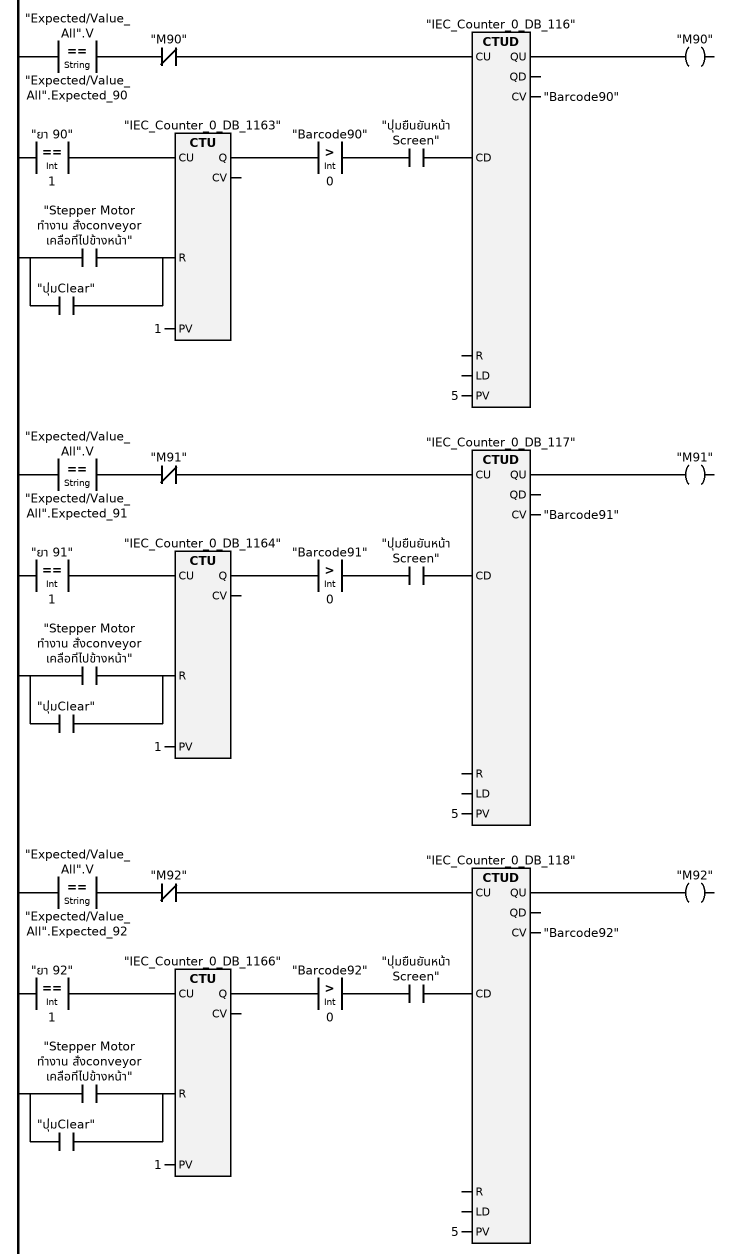
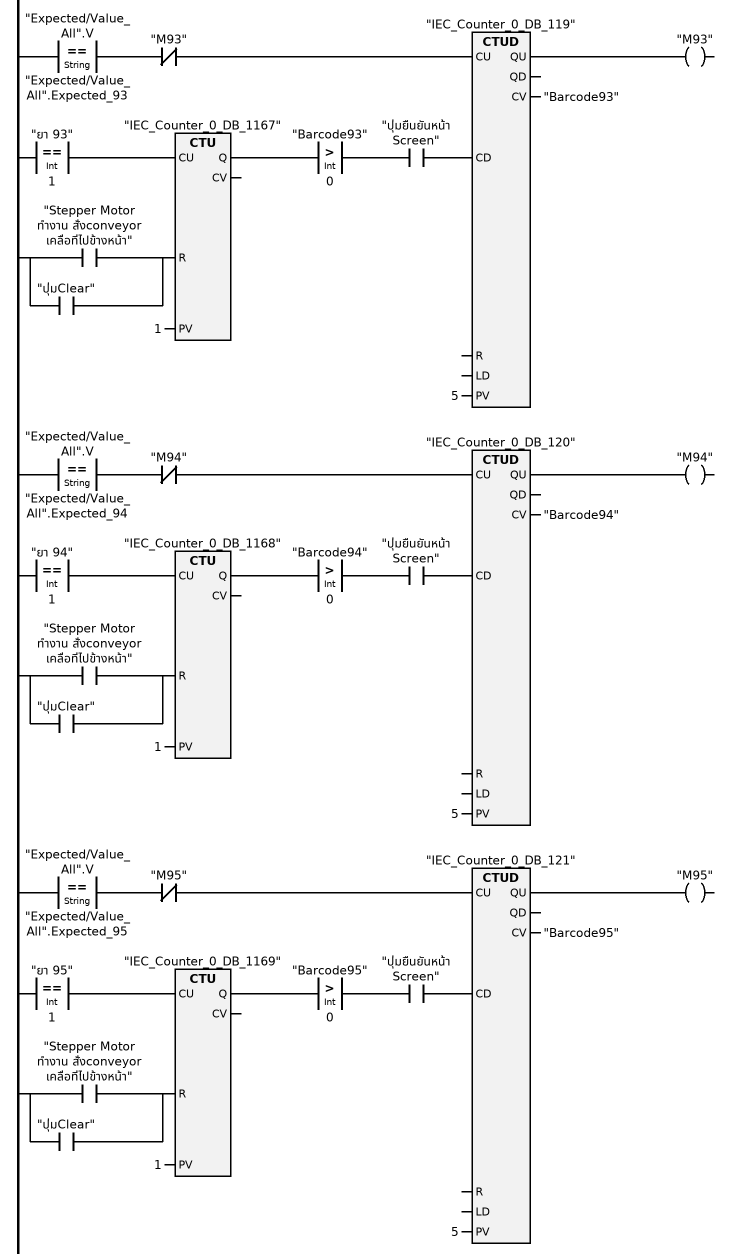
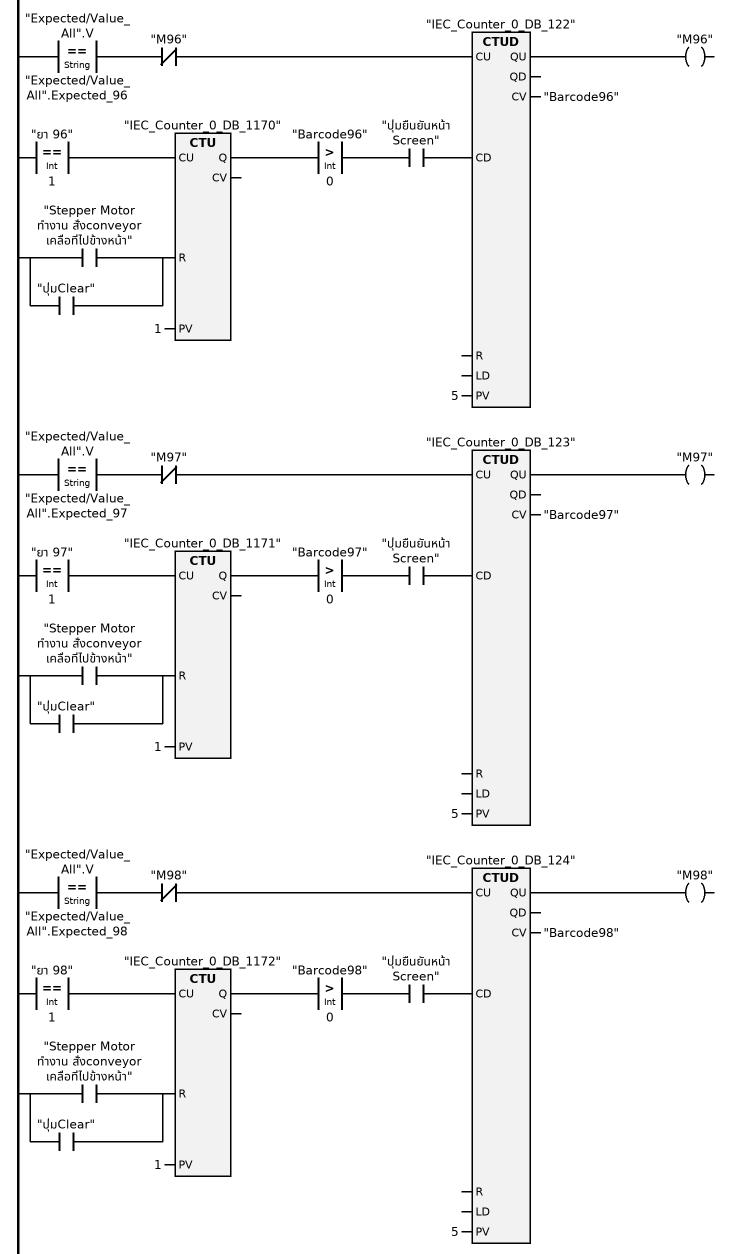
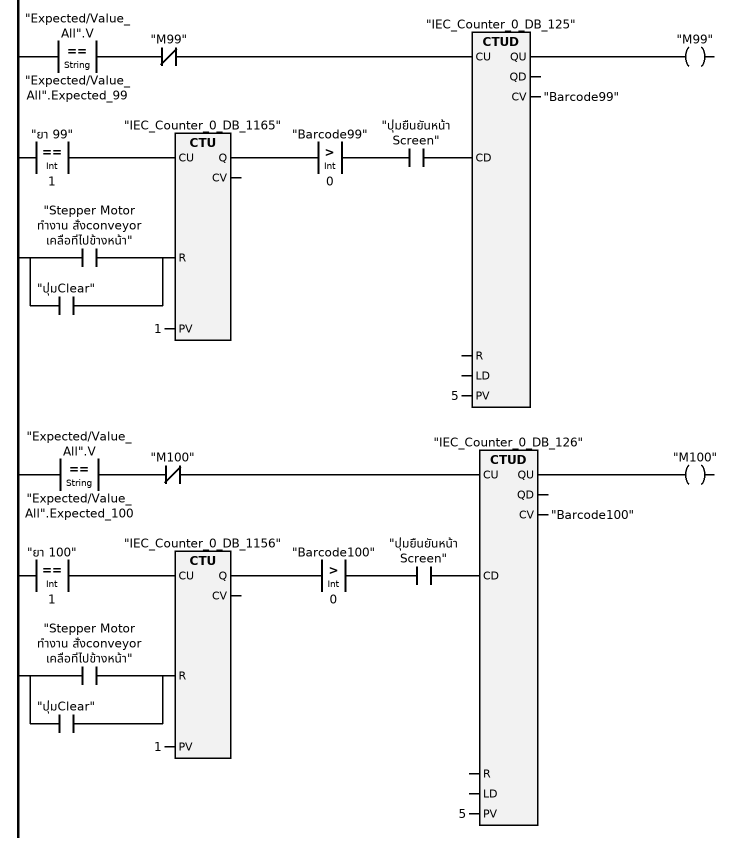
   "IEC_Counter_0_DB_1153".CTU(CU := "ยา 81" = 1,
                           R := "Stepper Motor ทำงาน สั่งconveyor เคลื่อที่ไปข้างหน้า" OR "ปุ่มClear",
                           PV := 1);
   "IEC_Counter_0_DB_107".CTUD(CU := ("Expected/Value_All".V = "Expected/Value_All".Expected_81) AND NOT "M81",
                           CD := "IEC_Counter_0_DB_1153".Q AND ("Barcode81" > 0) AND "ปุ่มยืนยันหน้า Screen",
                           PV := 5,
                           CV => "Barcode81");
   "M81" := "IEC_Counter_0_DB_107".QU;
   "IEC_Counter_0_DB_1154".CTU(CU := "ยา 82" = 1,
                           R := "Stepper Motor ทำงาน สั่งconveyor เคลื่อที่ไปข้างหน้า" OR "ปุ่มClear",
                           PV := 1);
   "IEC_Counter_0_DB_108".CTUD(CU := ("Expected/Value_All".V = "Expected/Value_All".Expected_82) AND NOT "M82",
                           CD := "IEC_Counter_0_DB_1154".Q AND ("Barcode82" > 0) AND "ปุ่มยืนยันหน้า Screen",
                           PV := 5,
                           CV => "Barcode82");
   "M82" := "IEC_Counter_0_DB_108".QU;
   "IEC_Counter_0_DB_1155".CTU(CU := "ยา 83" = 1,
                           R := "Stepper Motor ทำงาน สั่งconveyor เคลื่อที่ไปข้างหน้า" OR "ปุ่มClear",
                           PV := 1);
   "IEC_Counter_0_DB_109".CTUD(CU := ("Expected/Value_All".V = "Expected/Value_All".Expected_83) AND NOT "M83",
                           CD := "IEC_Counter_0_DB_1155".Q AND ("Barcode83" > 0) AND "ปุ่มยืนยันหน้า Screen",
                           PV := 5,
                           CV => "Barcode83");
   "M83" := "IEC_Counter_0_DB_109".QU;
   "IEC_Counter_0_DB_1157".CTU(CU := "ยา 84" = 1,
                           R := "Stepper Motor ทำงาน สั่งconveyor เคลื่อที่ไปข้างหน้า" OR "ปุ่มClear",
                           PV := 1);
   "IEC_Counter_0_DB_110".CTUD(CU := ("Expected/Value_All".V = "Expected/Value_All".Expected_84) AND NOT "M84",
                           CD := "IEC_Counter_0_DB_1157".Q AND ("Barcode84" > 0) AND "ปุ่มยืนยันหน้า Screen",
                           PV := 5,
                           CV => "Barcode84");
   "M84" := "IEC_Counter_0_DB_110".QU;
   "IEC_Counter_0_DB_1158".CTU(CU := "ยา 85" = 1,
                           R := "Stepper Motor ทำงาน สั่งconveyor เคลื่อที่ไปข้างหน้า" OR "ปุ่มClear",
                           PV := 1);
   "IEC_Counter_0_DB_111".CTUD(CU := ("Expected/Value_All".V = "Expected/Value_All".Expected_85) AND NOT "M85",
                           CD := "IEC_Counter_0_DB_1158".Q AND ("Barcode85" > 0) AND "ปุ่มยืนยันหน้า Screen",
                           PV := 5,
                           CV => "Barcode85");
   "M85" := "IEC_Counter_0_DB_111".QU;
   "IEC_Counter_0_DB_1159".CTU(CU := "ยา 86" = 1,
                           R := "Stepper Motor ทำงาน สั่งconveyor เคลื่อที่ไปข้างหน้า" OR "ปุ่มClear",
                           PV := 1);
   "IEC_Counter_0_DB_112".CTUD(CU := ("Expected/Value_All".V = "Expected/Value_All".Expected_86) AND NOT "M86",
                           CD := "IEC_Counter_0_DB_1159".Q AND ("Barcode86" > 0) AND "ปุ่มยืนยันหน้า Screen",
                           PV := 5,
                           CV => "Barcode86");
   "M86" := "IEC_Counter_0_DB_112".QU;
   "IEC_Counter_0_DB_1160".CTU(CU := "ยา 87" = 1,
                           R := "Stepper Motor ทำงาน สั่งconveyor เคลื่อที่ไปข้างหน้า" OR "ปุ่มClear",
                           PV := 1);
   "IEC_Counter_0_DB_113".CTUD(CU := ("Expected/Value_All".V = "Expected/Value_All".Expected_87) AND NOT "M87",
                           CD := "IEC_Counter_0_DB_1160".Q AND ("Barcode87" > 0) AND "ปุ่มยืนยันหน้า Screen",
                           PV := 5,
                           CV => "Barcode87");
   "M87" := "IEC_Counter_0_DB_113".QU;
   "IEC_Counter_0_DB_1161".CTU(CU := "ยา 88" = 1,
                           R := "Stepper Motor ทำงาน สั่งconveyor เคลื่อที่ไปข้างหน้า" OR "ปุ่มClear",
                           PV := 1);
   "IEC_Counter_0_DB_114".CTUD(CU := ("Expected/Value_All".V = "Expected/Value_All".Expected_88) AND NOT "M88",
                           CD := "IEC_Counter_0_DB_1161".Q AND ("Barcode88" > 0) AND "ปุ่มยืนยันหน้า Screen",
                           PV := 5,
                           CV => "Barcode88");
   "M88" := "IEC_Counter_0_DB_114".QU;
   "IEC_Counter_0_DB_1162".CTU(CU := "ยา 89" = 1,
                           R := "Stepper Motor ทำงาน สั่งconveyor เคลื่อที่ไปข้างหน้า" OR "ปุ่มClear",
                           PV := 1);
   "IEC_Counter_0_DB_115".CTUD(CU := ("Expected/Value_All".V = "Expected/Value_All".Expected_89) AND NOT "M89",
                           CD := "IEC_Counter_0_DB_1162".Q AND ("Barcode89" > 0) AND "ปุ่มยืนยันหน้า Screen",
                           PV := 5,
                           CV => "Barcode89");
   "M89" := "IEC_Counter_0_DB_115".QU;
   "IEC_Counter_0_DB_1163".CTU(CU := "ยา 90" = 1,
                           R := "Stepper Motor ทำงาน สั่งconveyor เคลื่อที่ไปข้างหน้า" OR "ปุ่มClear",
                           PV := 1);
   "IEC_Counter_0_DB_116".CTUD(CU := ("Expected/Value_All".V = "Expected/Value_All".Expected_90) AND NOT "M90",
                           CD := "IEC_Counter_0_DB_1163".Q AND ("Barcode90" > 0) AND "ปุ่มยืนยันหน้า Screen",
                           PV := 5,
                           CV => "Barcode90");
   "M90" := "IEC_Counter_0_DB_116".QU;
   "IEC_Counter_0_DB_1164".CTU(CU := "ยา 91" = 1,
                           R := "Stepper Motor ทำงาน สั่งconveyor เคลื่อที่ไปข้างหน้า" OR "ปุ่มClear",
                           PV := 1);
   "IEC_Counter_0_DB_117".CTUD(CU := ("Expected/Value_All".V = "Expected/Value_All".Expected_91) AND NOT "M91",
                           CD := "IEC_Counter_0_DB_1164".Q AND ("Barcode91" > 0) AND "ปุ่มยืนยันหน้า Screen",
                           PV := 5,
                           CV => "Barcode91");
   "M91" := "IEC_Counter_0_DB_117".QU;
   "IEC_Counter_0_DB_1166".CTU(CU := "ยา 92" = 1,
                           R := "Stepper Motor ทำงาน สั่งconveyor เคลื่อที่ไปข้างหน้า" OR "ปุ่มClear",
                           PV := 1);
   "IEC_Counter_0_DB_118".CTUD(CU := ("Expected/Value_All".V = "Expected/Value_All".Expected_92) AND NOT "M92",
                           CD := "IEC_Counter_0_DB_1166".Q AND ("Barcode92" > 0) AND "ปุ่มยืนยันหน้า Screen",
                           PV := 5,
                           CV => "Barcode92");
   "M92" := "IEC_Counter_0_DB_118".QU;
   "IEC_Counter_0_DB_1167".CTU(CU := "ยา 93" = 1,
                           R := "Stepper Motor ทำงาน สั่งconveyor เคลื่อที่ไปข้างหน้า" OR "ปุ่มClear",
                           PV := 1);
   "IEC_Counter_0_DB_119".CTUD(CU := ("Expected/Value_All".V = "Expected/Value_All".Expected_93) AND NOT "M93",
                           CD := "IEC_Counter_0_DB_1167".Q AND ("Barcode93" > 0) AND "ปุ่มยืนยันหน้า Screen",
                           PV := 5,
                           CV => "Barcode93");
   "M93" := "IEC_Counter_0_DB_119".QU;
   "IEC_Counter_0_DB_1168".CTU(CU := "ยา 94" = 1,
                           R := "Stepper Motor ทำงาน สั่งconveyor เคลื่อที่ไปข้างหน้า" OR "ปุ่มClear",
                           PV := 1);
   "IEC_Counter_0_DB_120".CTUD(CU := ("Expected/Value_All".V = "Expected/Value_All".Expected_94) AND NOT "M94",
                           CD := "IEC_Counter_0_DB_1168".Q AND ("Barcode94" > 0) AND "ปุ่มยืนยันหน้า Screen",
                           PV := 5,
                           CV => "Barcode94");
   "M94" := "IEC_Counter_0_DB_120".QU;
   "IEC_Counter_0_DB_1169".CTU(CU := "ยา 95" = 1,
                           R := "Stepper Motor ทำงาน สั่งconveyor เคลื่อที่ไปข้างหน้า" OR "ปุ่มClear",
                           PV := 1);
   "IEC_Counter_0_DB_121".CTUD(CU := ("Expected/Value_All".V = "Expected/Value_All".Expected_95) AND NOT "M95",
                           CD := "IEC_Counter_0_DB_1169".Q AND ("Barcode95" > 0) AND "ปุ่มยืนยันหน้า Screen",
                           PV := 5,
                           CV => "Barcode95");
   "M95" := "IEC_Counter_0_DB_121".QU;
   "IEC_Counter_0_DB_1170".CTU(CU := "ยา 96" = 1,
                           R := "Stepper Motor ทำงาน สั่งconveyor เคลื่อที่ไปข้างหน้า" OR "ปุ่มClear",
                           PV := 1);
   "IEC_Counter_0_DB_122".CTUD(CU := ("Expected/Value_All".V = "Expected/Value_All".Expected_96) AND NOT "M96",
                           CD := "IEC_Counter_0_DB_1170".Q AND ("Barcode96" > 0) AND "ปุ่มยืนยันหน้า Screen",
                           PV := 5,
                           CV => "Barcode96");
   "M96" := "IEC_Counter_0_DB_122".QU;
   "IEC_Counter_0_DB_1171".CTU(CU := "ยา 97" = 1,
                           R := "Stepper Motor ทำงาน สั่งconveyor เคลื่อที่ไปข้างหน้า" OR "ปุ่มClear",
                           PV := 1);
   "IEC_Counter_0_DB_123".CTUD(CU := ("Expected/Value_All".V = "Expected/Value_All".Expected_97) AND NOT "M97",
                           CD := "IEC_Counter_0_DB_1171".Q AND ("Barcode97" > 0) AND "ปุ่มยืนยันหน้า Screen",
                           PV := 5,
                           CV => "Barcode97");
   "M97" := "IEC_Counter_0_DB_123".QU;
   "IEC_Counter_0_DB_1172".CTU(CU := "ยา 98" = 1,
                           R := "Stepper Motor ทำงาน สั่งconveyor เคลื่อที่ไปข้างหน้า" OR "ปุ่มClear",
                           PV := 1);
   "IEC_Counter_0_DB_124".CTUD(CU := ("Expected/Value_All".V = "Expected/Value_All".Expected_98) AND NOT "M98",
                           CD := "IEC_Counter_0_DB_1172".Q AND ("Barcode98" > 0) AND "ปุ่มยืนยันหน้า Screen",
                           PV := 5,
                           CV => "Barcode98");
   "M98" := "IEC_Counter_0_DB_124".QU;
   "IEC_Counter_0_DB_1165".CTU(CU := "ยา 99" = 1,
                           R := "Stepper Motor ทำงาน สั่งconveyor เคลื่อที่ไปข้างหน้า" OR "ปุ่มClear",
                           PV := 1);
   "IEC_Counter_0_DB_125".CTUD(CU := ("Expected/Value_All".V = "Expected/Value_All".Expected_99) AND NOT "M99",
                           CD := "IEC_Counter_0_DB_1165".Q AND ("Barcode99" > 0) AND "ปุ่มยืนยันหน้า Screen",
                           PV := 5,
                           CV => "Barcode99");
   "M99" := "IEC_Counter_0_DB_125".QU;
   "IEC_Counter_0_DB_1156".CTU(CU := "ยา 100" = 1,
                           R := "Stepper Motor ทำงาน สั่งconveyor เคลื่อที่ไปข้างหน้า" OR "ปุ่มClear",
                           PV := 1);
   "IEC_Counter_0_DB_126".CTUD(CU := ("Expected/Value_All".V = "Expected/Value_All".Expected_100) AND NOT "M100",
                           CD := "IEC_Counter_0_DB_1156".Q AND ("Barcode100" > 0) AND "ปุ่มยืนยันหน้า Screen",
                           PV := 5,
                           CV => "Barcode100");
   "M100" := "IEC_Counter_0_DB_126".QU;
END_REGION

REGION Network 6
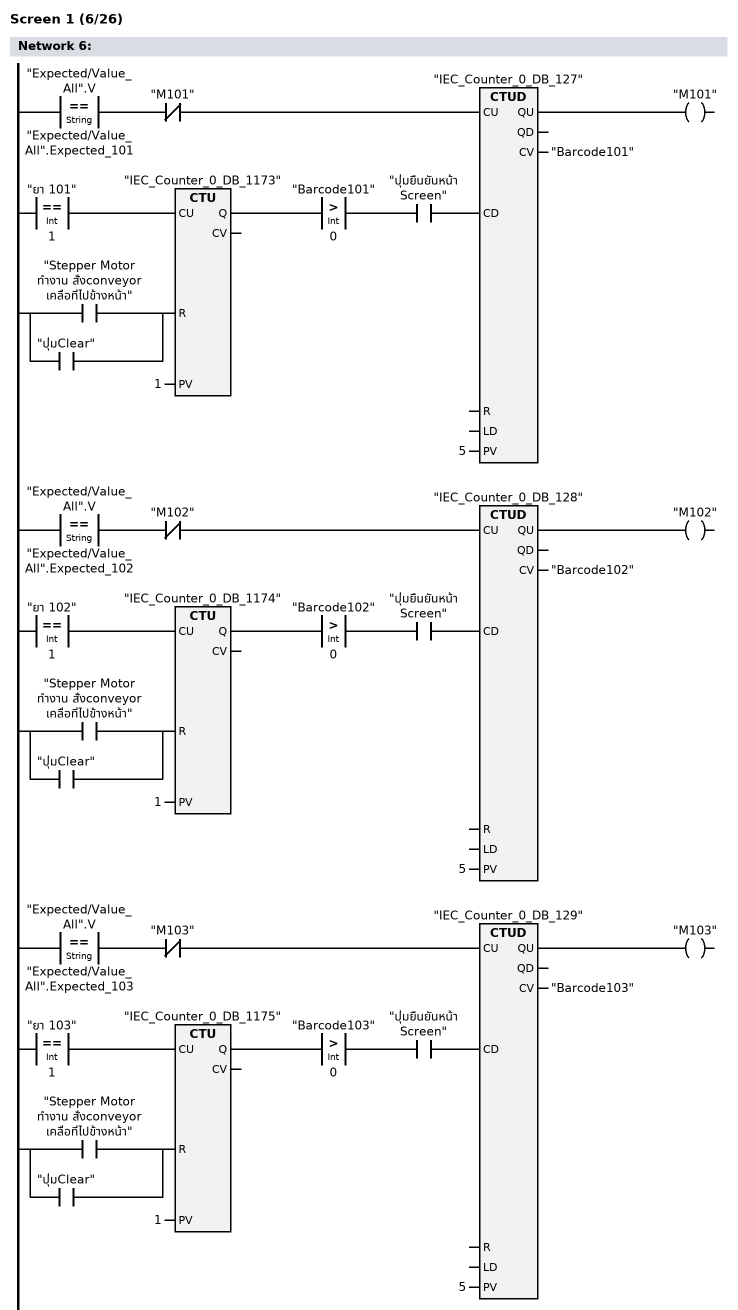
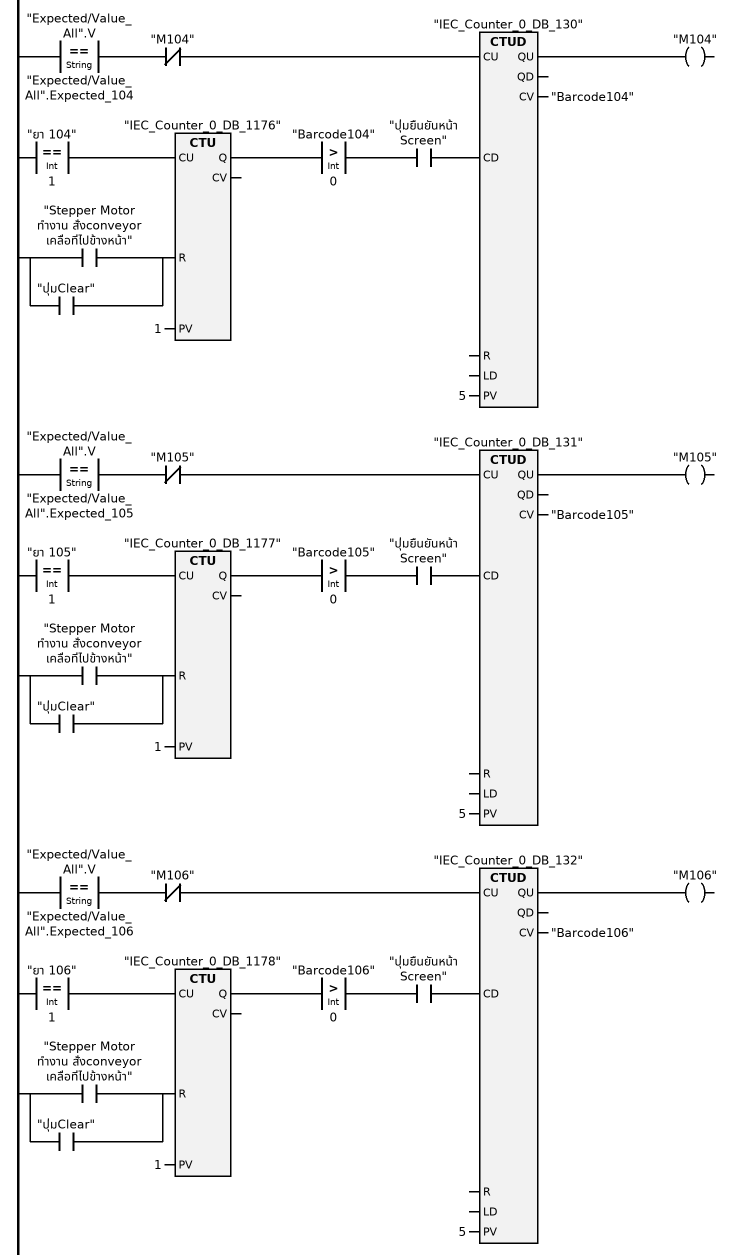
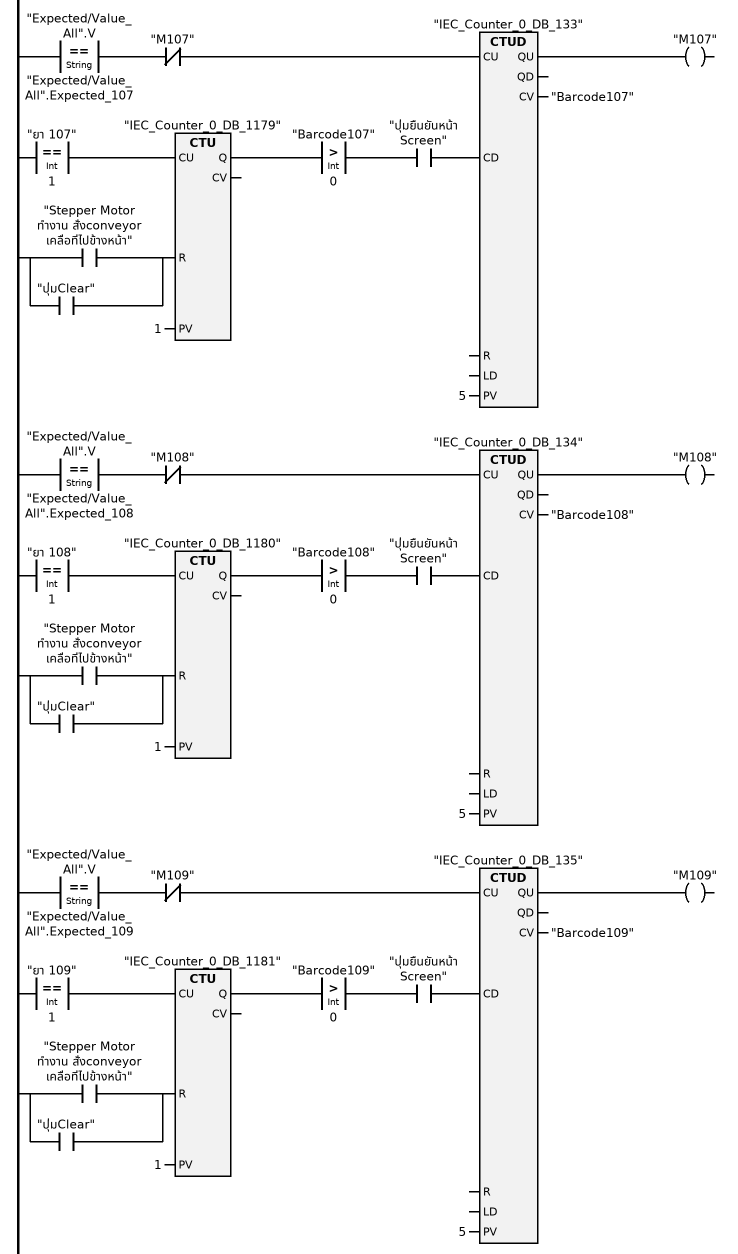
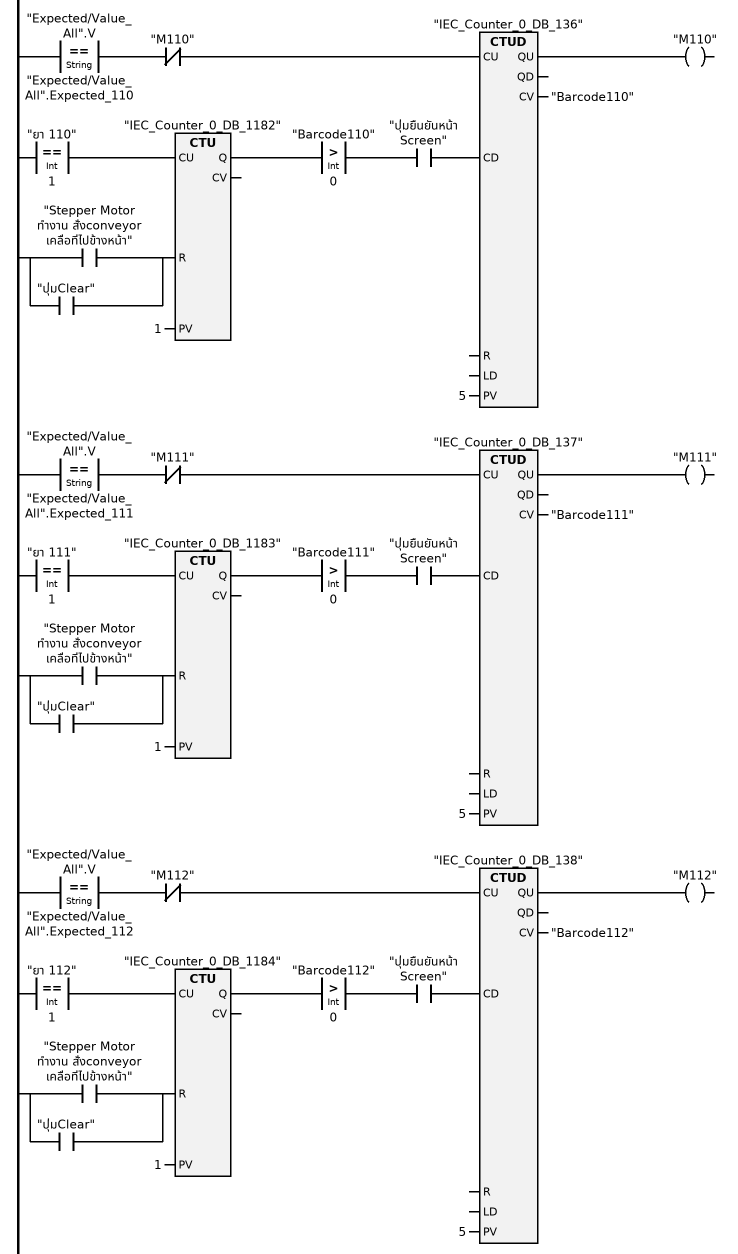
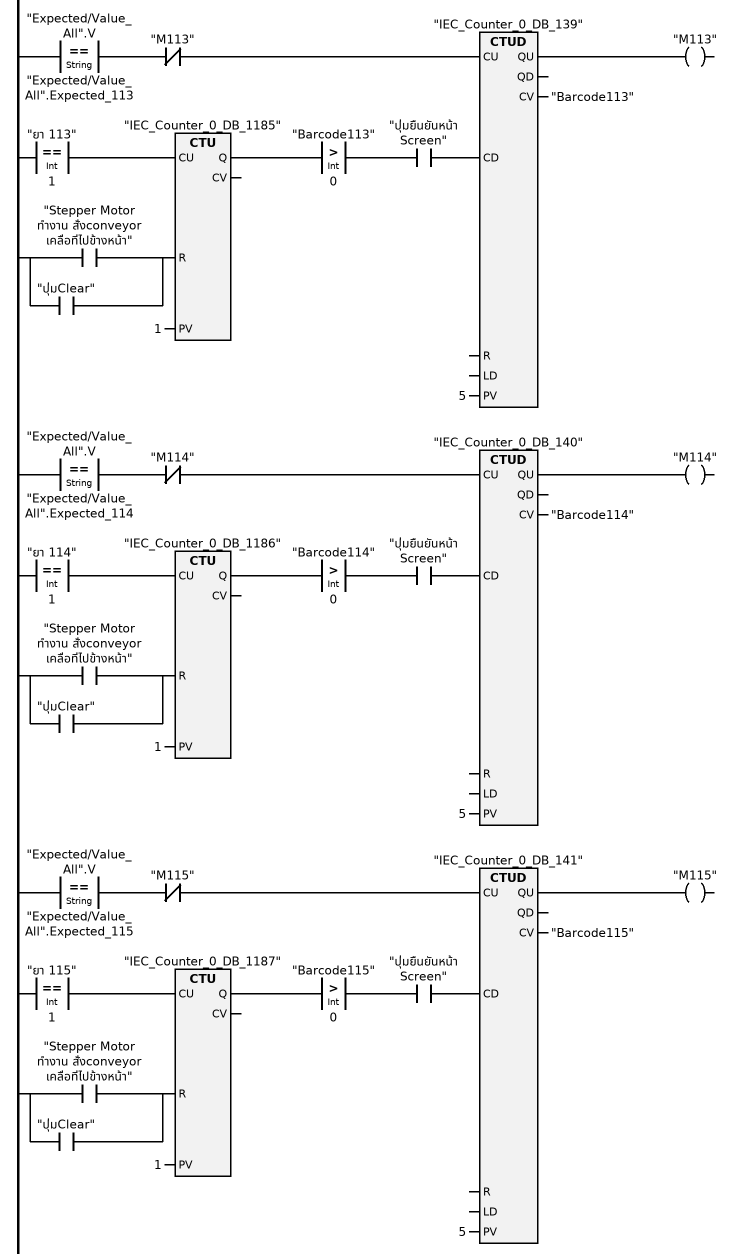
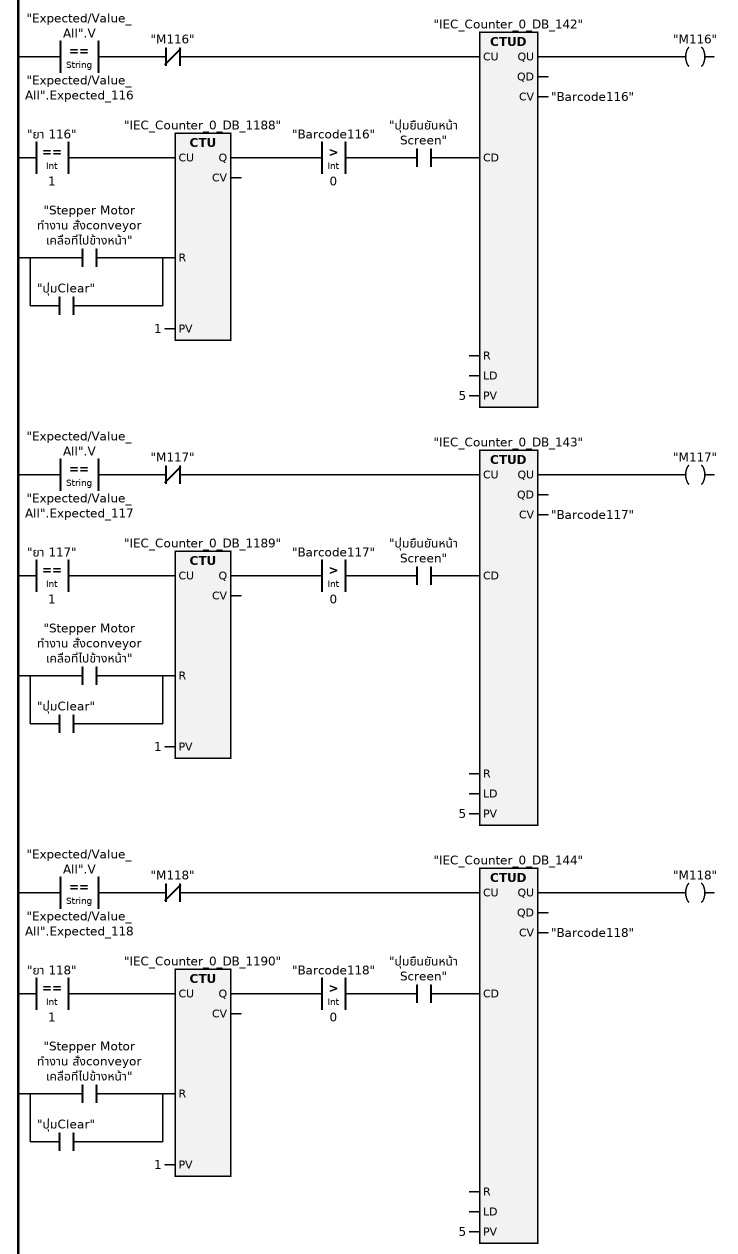
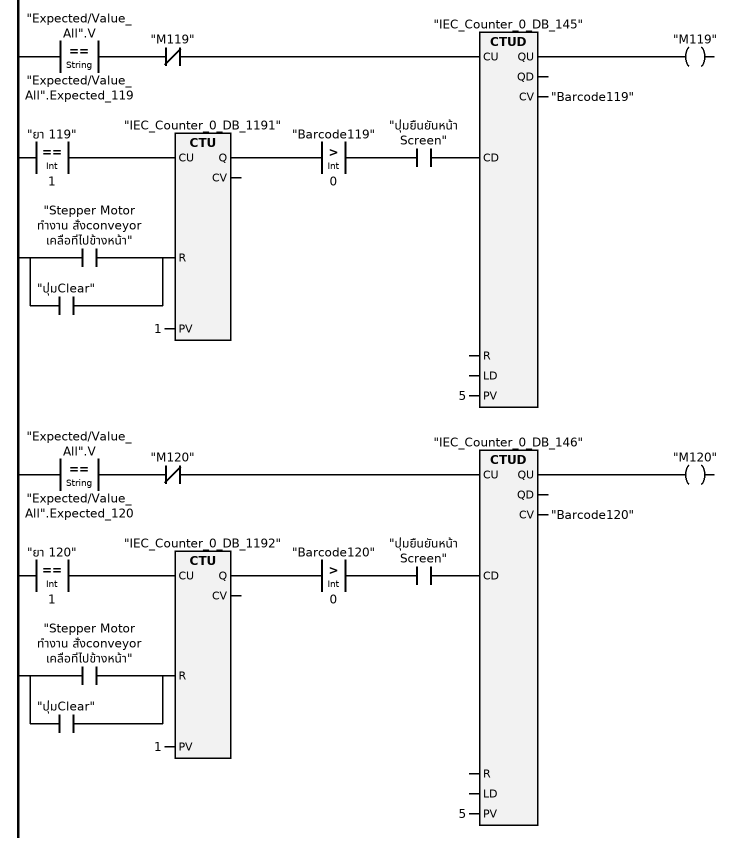
   "IEC_Counter_0_DB_1173".CTU(CU := "ยา 101" = 1,
                           R := "Stepper Motor ทำงาน สั่งconveyor เคลื่อที่ไปข้างหน้า" OR "ปุ่มClear",
                           PV := 1);
   "IEC_Counter_0_DB_127".CTUD(CU := ("Expected/Value_All".V = "Expected/Value_All".Expected_101) AND NOT "M101",
                           CD := "IEC_Counter_0_DB_1173".Q AND ("Barcode101" > 0) AND "ปุ่มยืนยันหน้า Screen",
                           PV := 5,
                           CV => "Barcode101");
   "M101" := "IEC_Counter_0_DB_127".QU;
   "IEC_Counter_0_DB_1174".CTU(CU := "ยา 102" = 1,
                           R := "Stepper Motor ทำงาน สั่งconveyor เคลื่อที่ไปข้างหน้า" OR "ปุ่มClear",
                           PV := 1);
   "IEC_Counter_0_DB_128".CTUD(CU := ("Expected/Value_All".V = "Expected/Value_All".Expected_102) AND NOT "M102",
                           CD := "IEC_Counter_0_DB_1174".Q AND ("Barcode102" > 0) AND "ปุ่มยืนยันหน้า Screen",
                           PV := 5,
                           CV => "Barcode102");
   "M102" := "IEC_Counter_0_DB_128".QU;
   "IEC_Counter_0_DB_1175".CTU(CU := "ยา 103" = 1,
                           R := "Stepper Motor ทำงาน สั่งconveyor เคลื่อที่ไปข้างหน้า" OR "ปุ่มClear",
                           PV := 1);
   "IEC_Counter_0_DB_129".CTUD(CU := ("Expected/Value_All".V = "Expected/Value_All".Expected_103) AND NOT "M103",
                           CD := "IEC_Counter_0_DB_1175".Q AND ("Barcode103" > 0) AND "ปุ่มยืนยันหน้า Screen",
                           PV := 5,
                           CV => "Barcode103");
   "M103" := "IEC_Counter_0_DB_129".QU;
   "IEC_Counter_0_DB_1176".CTU(CU := "ยา 104" = 1,
                           R := "Stepper Motor ทำงาน สั่งconveyor เคลื่อที่ไปข้างหน้า" OR "ปุ่มClear",
                           PV := 1);
   "IEC_Counter_0_DB_130".CTUD(CU := ("Expected/Value_All".V = "Expected/Value_All".Expected_104) AND NOT "M104",
                           CD := "IEC_Counter_0_DB_1176".Q AND ("Barcode104" > 0) AND "ปุ่มยืนยันหน้า Screen",
                           PV := 5,
                           CV => "Barcode104");
   "M104" := "IEC_Counter_0_DB_130".QU;
   "IEC_Counter_0_DB_1177".CTU(CU := "ยา 105" = 1,
                           R := "Stepper Motor ทำงาน สั่งconveyor เคลื่อที่ไปข้างหน้า" OR "ปุ่มClear",
                           PV := 1);
   "IEC_Counter_0_DB_131".CTUD(CU := ("Expected/Value_All".V = "Expected/Value_All".Expected_105) AND NOT "M105",
                           CD := "IEC_Counter_0_DB_1177".Q AND ("Barcode105" > 0) AND "ปุ่มยืนยันหน้า Screen",
                           PV := 5,
                           CV => "Barcode105");
   "M105" := "IEC_Counter_0_DB_131".QU;
   "IEC_Counter_0_DB_1178".CTU(CU := "ยา 106" = 1,
                           R := "Stepper Motor ทำงาน สั่งconveyor เคลื่อที่ไปข้างหน้า" OR "ปุ่มClear",
                           PV := 1);
   "IEC_Counter_0_DB_132".CTUD(CU := ("Expected/Value_All".V = "Expected/Value_All".Expected_106) AND NOT "M106",
                           CD := "IEC_Counter_0_DB_1178".Q AND ("Barcode106" > 0) AND "ปุ่มยืนยันหน้า Screen",
                           PV := 5,
                           CV => "Barcode106");
   "M106" := "IEC_Counter_0_DB_132".QU;
   "IEC_Counter_0_DB_1179".CTU(CU := "ยา 107" = 1,
                           R := "Stepper Motor ทำงาน สั่งconveyor เคลื่อที่ไปข้างหน้า" OR "ปุ่มClear",
                           PV := 1);
   "IEC_Counter_0_DB_133".CTUD(CU := ("Expected/Value_All".V = "Expected/Value_All".Expected_107) AND NOT "M107",
                           CD := "IEC_Counter_0_DB_1179".Q AND ("Barcode107" > 0) AND "ปุ่มยืนยันหน้า Screen",
                           PV := 5,
                           CV => "Barcode107");
   "M107" := "IEC_Counter_0_DB_133".QU;
   "IEC_Counter_0_DB_1180".CTU(CU := "ยา 108" = 1,
                           R := "Stepper Motor ทำงาน สั่งconveyor เคลื่อที่ไปข้างหน้า" OR "ปุ่มClear",
                           PV := 1);
   "IEC_Counter_0_DB_134".CTUD(CU := ("Expected/Value_All".V = "Expected/Value_All".Expected_108) AND NOT "M108",
                           CD := "IEC_Counter_0_DB_1180".Q AND ("Barcode108" > 0) AND "ปุ่มยืนยันหน้า Screen",
                           PV := 5,
                           CV => "Barcode108");
   "M108" := "IEC_Counter_0_DB_134".QU;
   "IEC_Counter_0_DB_1181".CTU(CU := "ยา 109" = 1,
                           R := "Stepper Motor ทำงาน สั่งconveyor เคลื่อที่ไปข้างหน้า" OR "ปุ่มClear",
                           PV := 1);
   "IEC_Counter_0_DB_135".CTUD(CU := ("Expected/Value_All".V = "Expected/Value_All".Expected_109) AND NOT "M109",
                           CD := "IEC_Counter_0_DB_1181".Q AND ("Barcode109" > 0) AND "ปุ่มยืนยันหน้า Screen",
                           PV := 5,
                           CV => "Barcode109");
   "M109" := "IEC_Counter_0_DB_135".QU;
   "IEC_Counter_0_DB_1182".CTU(CU := "ยา 110" = 1,
                           R := "Stepper Motor ทำงาน สั่งconveyor เคลื่อที่ไปข้างหน้า" OR "ปุ่มClear",
                           PV := 1);
   "IEC_Counter_0_DB_136".CTUD(CU := ("Expected/Value_All".V = "Expected/Value_All".Expected_110) AND NOT "M110",
                           CD := "IEC_Counter_0_DB_1182".Q AND ("Barcode110" > 0) AND "ปุ่มยืนยันหน้า Screen",
                           PV := 5,
                           CV => "Barcode110");
   "M110" := "IEC_Counter_0_DB_136".QU;
   "IEC_Counter_0_DB_1183".CTU(CU := "ยา 111" = 1,
                           R := "Stepper Motor ทำงาน สั่งconveyor เคลื่อที่ไปข้างหน้า" OR "ปุ่มClear",
                           PV := 1);
   "IEC_Counter_0_DB_137".CTUD(CU := ("Expected/Value_All".V = "Expected/Value_All".Expected_111) AND NOT "M111",
                           CD := "IEC_Counter_0_DB_1183".Q AND ("Barcode111" > 0) AND "ปุ่มยืนยันหน้า Screen",
                           PV := 5,
                           CV => "Barcode111");
   "M111" := "IEC_Counter_0_DB_137".QU;
   "IEC_Counter_0_DB_1184".CTU(CU := "ยา 112" = 1,
                           R := "Stepper Motor ทำงาน สั่งconveyor เคลื่อที่ไปข้างหน้า" OR "ปุ่มClear",
                           PV := 1);
   "IEC_Counter_0_DB_138".CTUD(CU := ("Expected/Value_All".V = "Expected/Value_All".Expected_112) AND NOT "M112",
                           CD := "IEC_Counter_0_DB_1184".Q AND ("Barcode112" > 0) AND "ปุ่มยืนยันหน้า Screen",
                           PV := 5,
                           CV => "Barcode112");
   "M112" := "IEC_Counter_0_DB_138".QU;
   "IEC_Counter_0_DB_1185".CTU(CU := "ยา 113" = 1,
                           R := "Stepper Motor ทำงาน สั่งconveyor เคลื่อที่ไปข้างหน้า" OR "ปุ่มClear",
                           PV := 1);
   "IEC_Counter_0_DB_139".CTUD(CU := ("Expected/Value_All".V = "Expected/Value_All".Expected_113) AND NOT "M113",
                           CD := "IEC_Counter_0_DB_1185".Q AND ("Barcode113" > 0) AND "ปุ่มยืนยันหน้า Screen",
                           PV := 5,
                           CV => "Barcode113");
   "M113" := "IEC_Counter_0_DB_139".QU;
   "IEC_Counter_0_DB_1186".CTU(CU := "ยา 114" = 1,
                           R := "Stepper Motor ทำงาน สั่งconveyor เคลื่อที่ไปข้างหน้า" OR "ปุ่มClear",
                           PV := 1);
   "IEC_Counter_0_DB_140".CTUD(CU := ("Expected/Value_All".V = "Expected/Value_All".Expected_114) AND NOT "M114",
                           CD := "IEC_Counter_0_DB_1186".Q AND ("Barcode114" > 0) AND "ปุ่มยืนยันหน้า Screen",
                           PV := 5,
                           CV => "Barcode114");
   "M114" := "IEC_Counter_0_DB_140".QU;
   "IEC_Counter_0_DB_1187".CTU(CU := "ยา 115" = 1,
                           R := "Stepper Motor ทำงาน สั่งconveyor เคลื่อที่ไปข้างหน้า" OR "ปุ่มClear",
                           PV := 1);
   "IEC_Counter_0_DB_141".CTUD(CU := ("Expected/Value_All".V = "Expected/Value_All".Expected_115) AND NOT "M115",
                           CD := "IEC_Counter_0_DB_1187".Q AND ("Barcode115" > 0) AND "ปุ่มยืนยันหน้า Screen",
                           PV := 5,
                           CV => "Barcode115");
   "M115" := "IEC_Counter_0_DB_141".QU;
   "IEC_Counter_0_DB_1188".CTU(CU := "ยา 116" = 1,
                           R := "Stepper Motor ทำงาน สั่งconveyor เคลื่อที่ไปข้างหน้า" OR "ปุ่มClear",
                           PV := 1);
   "IEC_Counter_0_DB_142".CTUD(CU := ("Expected/Value_All".V = "Expected/Value_All".Expected_116) AND NOT "M116",
                           CD := "IEC_Counter_0_DB_1188".Q AND ("Barcode116" > 0) AND "ปุ่มยืนยันหน้า Screen",
                           PV := 5,
                           CV => "Barcode116");
   "M116" := "IEC_Counter_0_DB_142".QU;
   "IEC_Counter_0_DB_1189".CTU(CU := "ยา 117" = 1,
                           R := "Stepper Motor ทำงาน สั่งconveyor เคลื่อที่ไปข้างหน้า" OR "ปุ่มClear",
                           PV := 1);
   "IEC_Counter_0_DB_143".CTUD(CU := ("Expected/Value_All".V = "Expected/Value_All".Expected_117) AND NOT "M117",
                           CD := "IEC_Counter_0_DB_1189".Q AND ("Barcode117" > 0) AND "ปุ่มยืนยันหน้า Screen",
                           PV := 5,
                           CV => "Barcode117");
   "M117" := "IEC_Counter_0_DB_143".QU;
   "IEC_Counter_0_DB_1190".CTU(CU := "ยา 118" = 1,
                           R := "Stepper Motor ทำงาน สั่งconveyor เคลื่อที่ไปข้างหน้า" OR "ปุ่มClear",
                           PV := 1);
   "IEC_Counter_0_DB_144".CTUD(CU := ("Expected/Value_All".V = "Expected/Value_All".Expected_118) AND NOT "M118",
                           CD := "IEC_Counter_0_DB_1190".Q AND ("Barcode118" > 0) AND "ปุ่มยืนยันหน้า Screen",
                           PV := 5,
                           CV => "Barcode118");
   "M118" := "IEC_Counter_0_DB_144".QU;
   "IEC_Counter_0_DB_1191".CTU(CU := "ยา 119" = 1,
                           R := "Stepper Motor ทำงาน สั่งconveyor เคลื่อที่ไปข้างหน้า" OR "ปุ่มClear",
                           PV := 1);
   "IEC_Counter_0_DB_145".CTUD(CU := ("Expected/Value_All".V = "Expected/Value_All".Expected_119) AND NOT "M119",
                           CD := "IEC_Counter_0_DB_1191".Q AND ("Barcode119" > 0) AND "ปุ่มยืนยันหน้า Screen",
                           PV := 5,
                           CV => "Barcode119");
   "M119" := "IEC_Counter_0_DB_145".QU;
   "IEC_Counter_0_DB_1192".CTU(CU := "ยา 120" = 1,
                           R := "Stepper Motor ทำงาน สั่งconveyor เคลื่อที่ไปข้างหน้า" OR "ปุ่มClear",
                           PV := 1);
   "IEC_Counter_0_DB_146".CTUD(CU := ("Expected/Value_All".V = "Expected/Value_All".Expected_120) AND NOT "M120",
                           CD := "IEC_Counter_0_DB_1192".Q AND ("Barcode120" > 0) AND "ปุ่มยืนยันหน้า Screen",
                           PV := 5,
                           CV => "Barcode120");
   "M120" := "IEC_Counter_0_DB_146".QU;
END_REGION

REGION Network 7
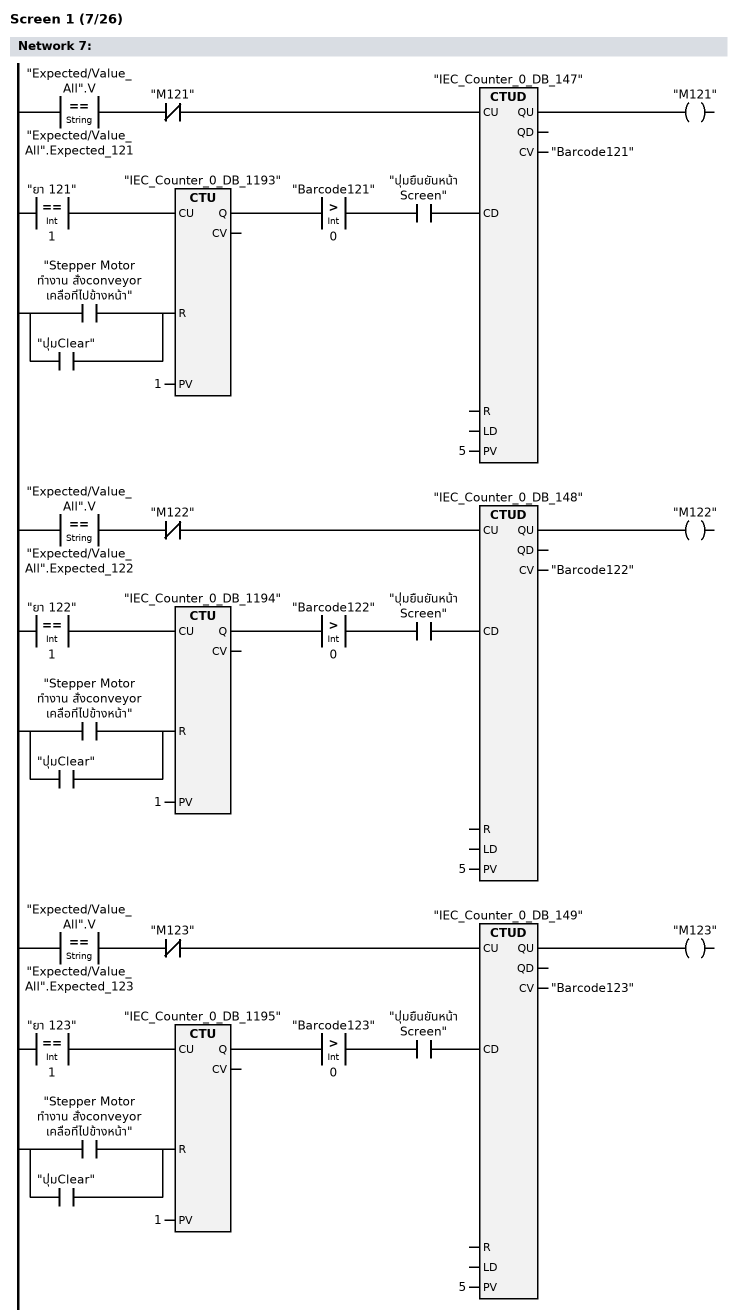
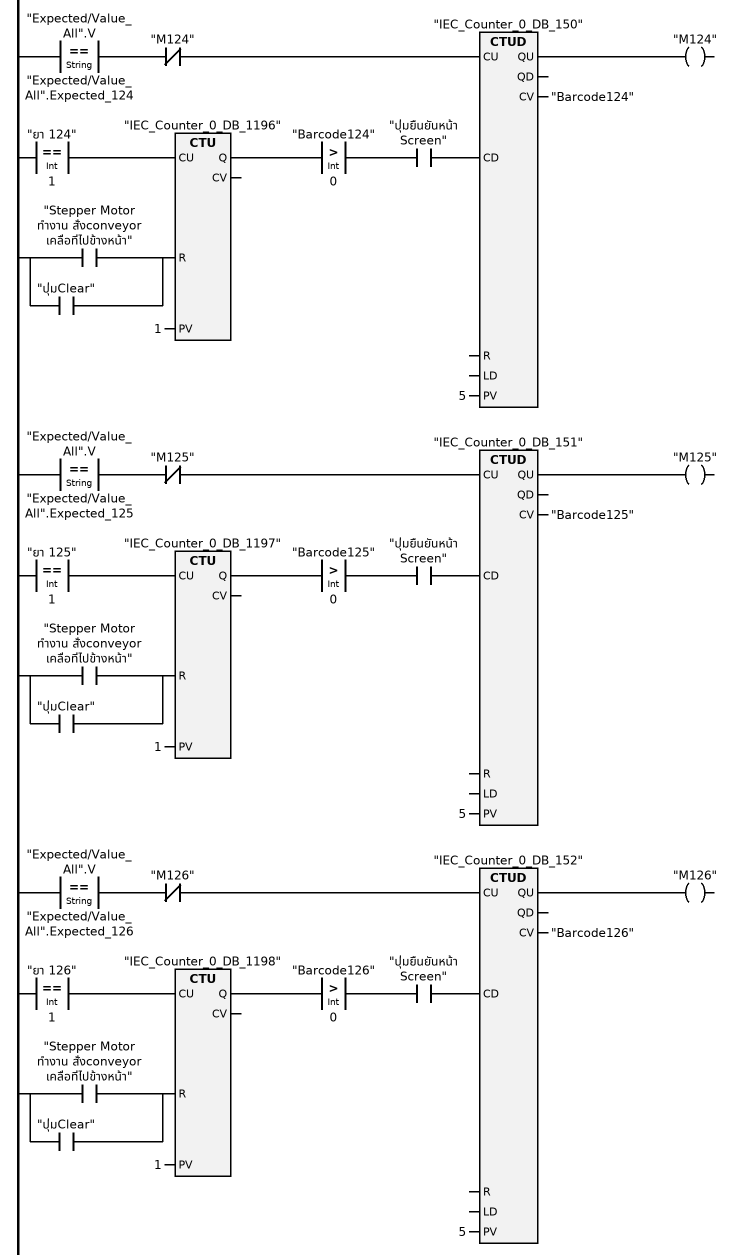
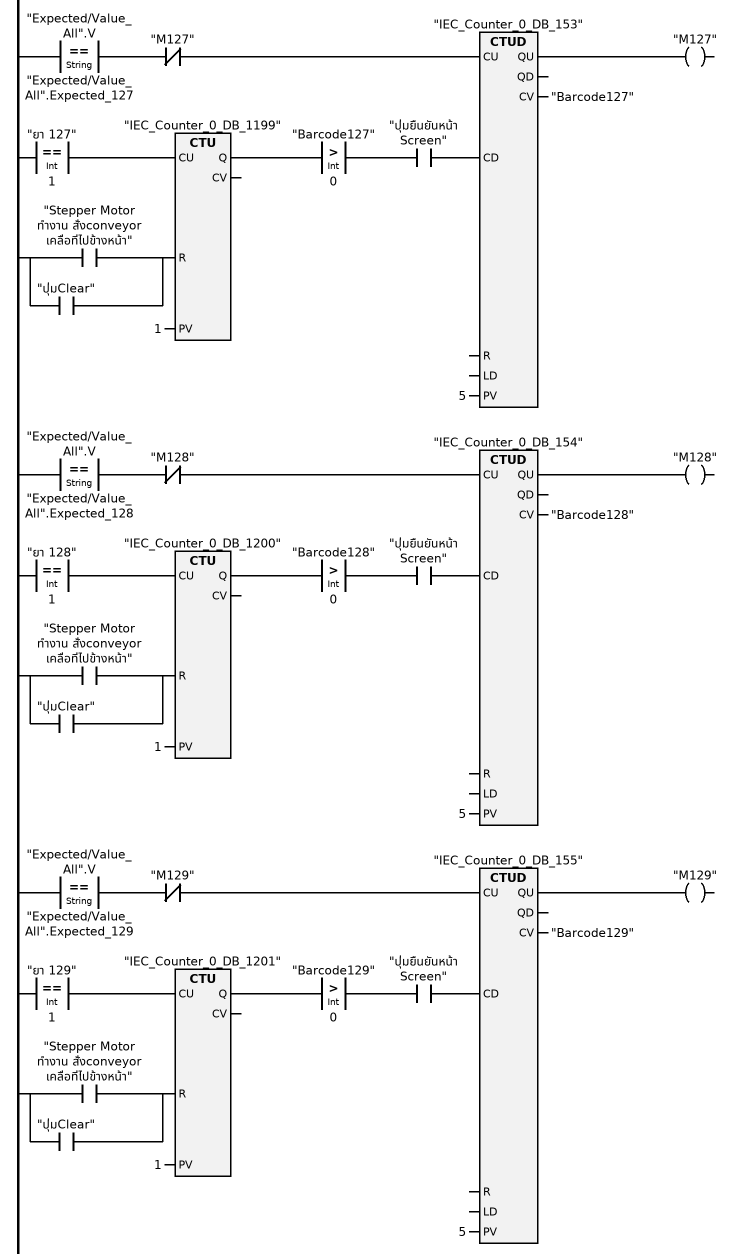
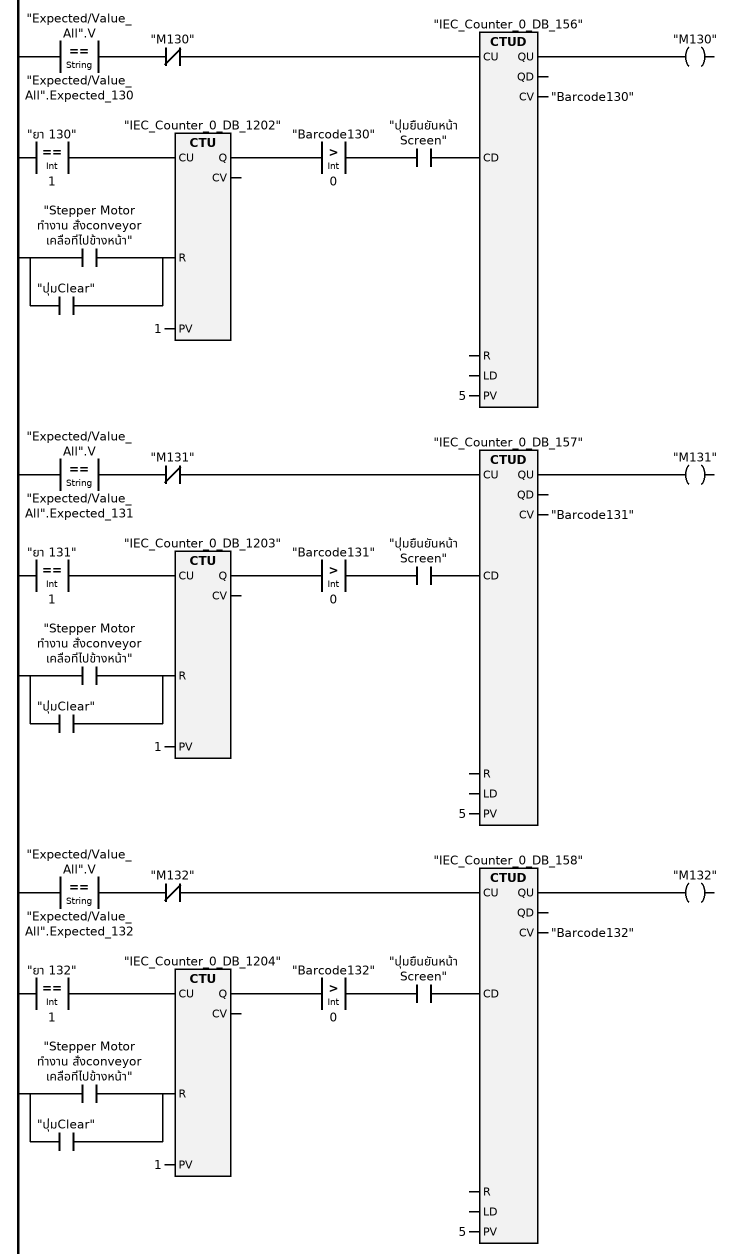
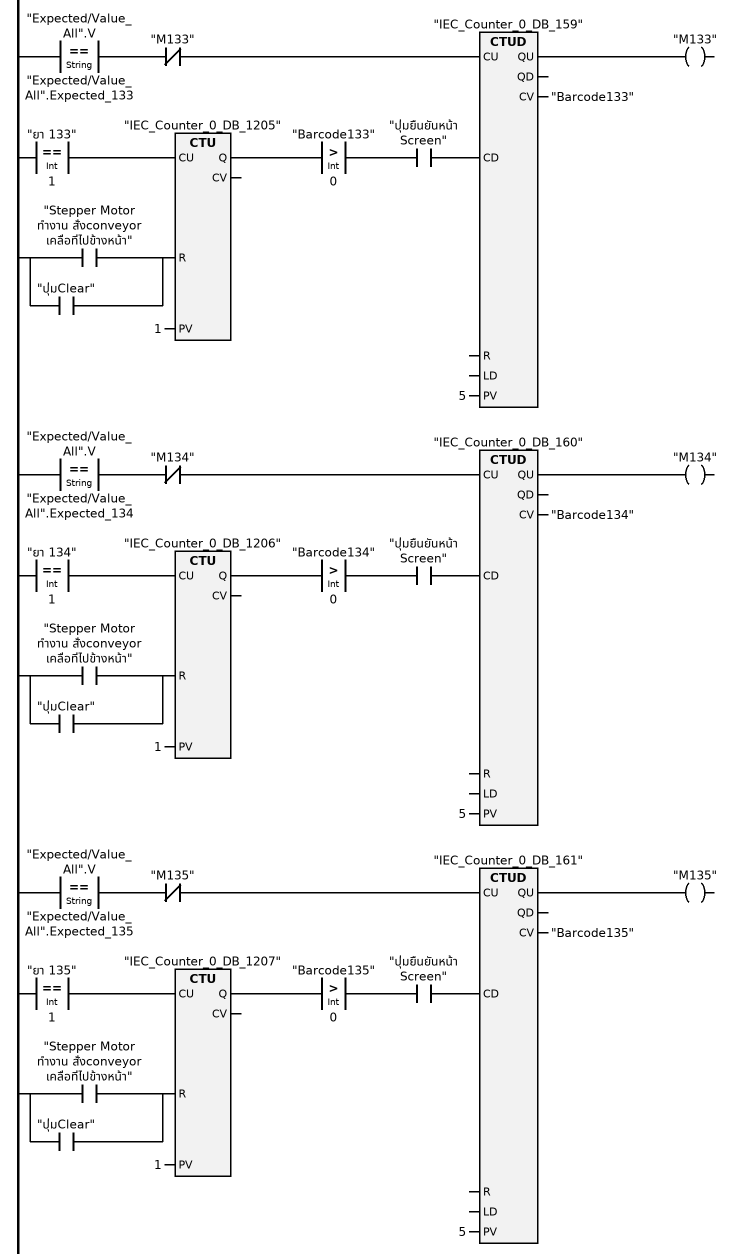
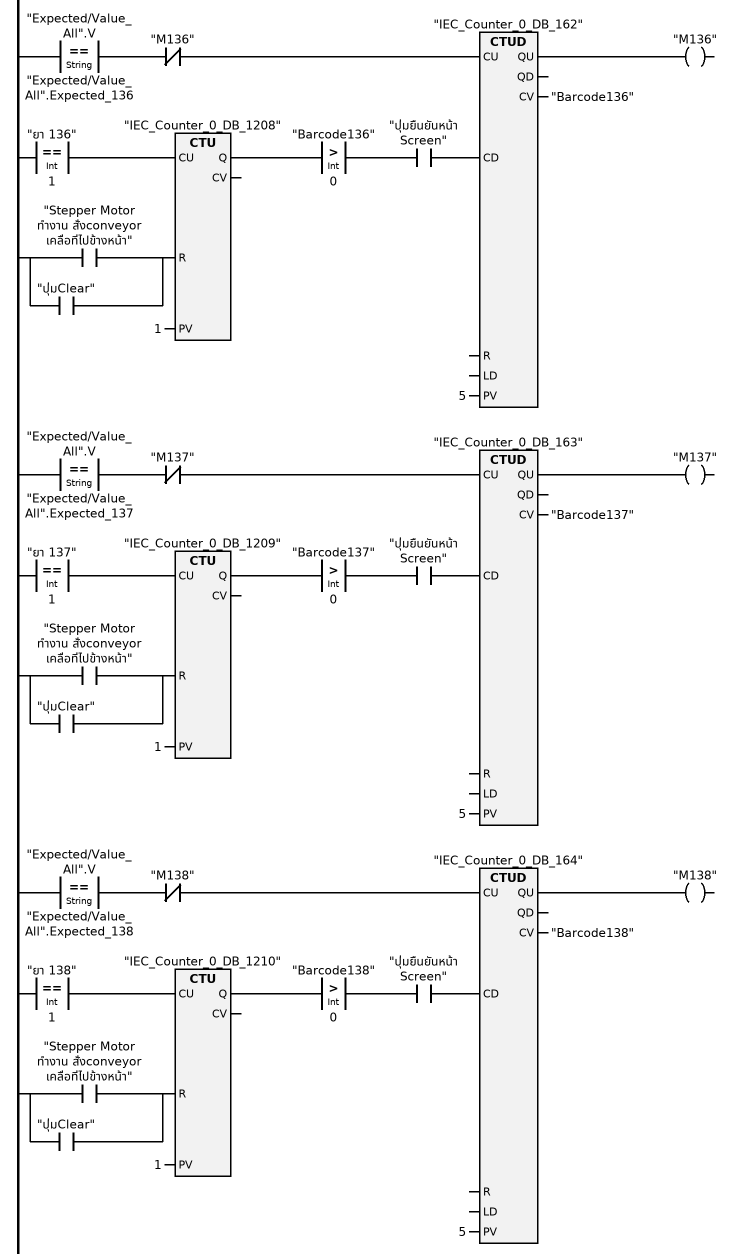
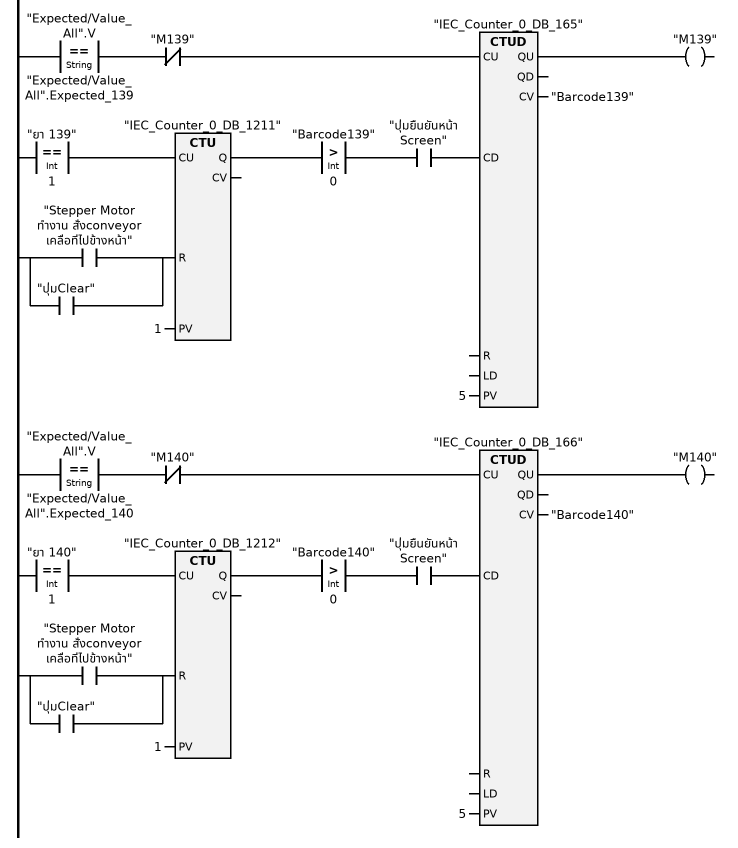
   "IEC_Counter_0_DB_1193".CTU(CU := "ยา 121" = 1,
                           R := "Stepper Motor ทำงาน สั่งconveyor เคลื่อที่ไปข้างหน้า" OR "ปุ่มClear",
                           PV := 1);
   "IEC_Counter_0_DB_147".CTUD(CU := ("Expected/Value_All".V = "Expected/Value_All".Expected_121) AND NOT "M121",
                           CD := "IEC_Counter_0_DB_1193".Q AND ("Barcode121" > 0) AND "ปุ่มยืนยันหน้า Screen",
                           PV := 5,
                           CV => "Barcode121");
   "M121" := "IEC_Counter_0_DB_147".QU;
   "IEC_Counter_0_DB_1194".CTU(CU := "ยา 122" = 1,
                           R := "Stepper Motor ทำงาน สั่งconveyor เคลื่อที่ไปข้างหน้า" OR "ปุ่มClear",
                           PV := 1);
   "IEC_Counter_0_DB_148".CTUD(CU := ("Expected/Value_All".V = "Expected/Value_All".Expected_122) AND NOT "M122",
                           CD := "IEC_Counter_0_DB_1194".Q AND ("Barcode122" > 0) AND "ปุ่มยืนยันหน้า Screen",
                           PV := 5,
                           CV => "Barcode122");
   "M122" := "IEC_Counter_0_DB_148".QU;
   "IEC_Counter_0_DB_1195".CTU(CU := "ยา 123" = 1,
                           R := "Stepper Motor ทำงาน สั่งconveyor เคลื่อที่ไปข้างหน้า" OR "ปุ่มClear",
                           PV := 1);
   "IEC_Counter_0_DB_149".CTUD(CU := ("Expected/Value_All".V = "Expected/Value_All".Expected_123) AND NOT "M123",
                           CD := "IEC_Counter_0_DB_1195".Q AND ("Barcode123" > 0) AND "ปุ่มยืนยันหน้า Screen",
                           PV := 5,
                           CV => "Barcode123");
   "M123" := "IEC_Counter_0_DB_149".QU;
   "IEC_Counter_0_DB_1196".CTU(CU := "ยา 124" = 1,
                           R := "Stepper Motor ทำงาน สั่งconveyor เคลื่อที่ไปข้างหน้า" OR "ปุ่มClear",
                           PV := 1);
   "IEC_Counter_0_DB_150".CTUD(CU := ("Expected/Value_All".V = "Expected/Value_All".Expected_124) AND NOT "M124",
                           CD := "IEC_Counter_0_DB_1196".Q AND ("Barcode124" > 0) AND "ปุ่มยืนยันหน้า Screen",
                           PV := 5,
                           CV => "Barcode124");
   "M124" := "IEC_Counter_0_DB_150".QU;
   "IEC_Counter_0_DB_1197".CTU(CU := "ยา 125" = 1,
                           R := "Stepper Motor ทำงาน สั่งconveyor เคลื่อที่ไปข้างหน้า" OR "ปุ่มClear",
                           PV := 1);
   "IEC_Counter_0_DB_151".CTUD(CU := ("Expected/Value_All".V = "Expected/Value_All".Expected_125) AND NOT "M125",
                           CD := "IEC_Counter_0_DB_1197".Q AND ("Barcode125" > 0) AND "ปุ่มยืนยันหน้า Screen",
                           PV := 5,
                           CV => "Barcode125");
   "M125" := "IEC_Counter_0_DB_151".QU;
   "IEC_Counter_0_DB_1198".CTU(CU := "ยา 126" = 1,
                           R := "Stepper Motor ทำงาน สั่งconveyor เคลื่อที่ไปข้างหน้า" OR "ปุ่มClear",
                           PV := 1);
   "IEC_Counter_0_DB_152".CTUD(CU := ("Expected/Value_All".V = "Expected/Value_All".Expected_126) AND NOT "M126",
                           CD := "IEC_Counter_0_DB_1198".Q AND ("Barcode126" > 0) AND "ปุ่มยืนยันหน้า Screen",
                           PV := 5,
                           CV => "Barcode126");
   "M126" := "IEC_Counter_0_DB_152".QU;
   "IEC_Counter_0_DB_1199".CTU(CU := "ยา 127" = 1,
                           R := "Stepper Motor ทำงาน สั่งconveyor เคลื่อที่ไปข้างหน้า" OR "ปุ่มClear",
                           PV := 1);
   "IEC_Counter_0_DB_153".CTUD(CU := ("Expected/Value_All".V = "Expected/Value_All".Expected_127) AND NOT "M127",
                           CD := "IEC_Counter_0_DB_1199".Q AND ("Barcode127" > 0) AND "ปุ่มยืนยันหน้า Screen",
                           PV := 5,
                           CV => "Barcode127");
   "M127" := "IEC_Counter_0_DB_153".QU;
   "IEC_Counter_0_DB_1200".CTU(CU := "ยา 128" = 1,
                           R := "Stepper Motor ทำงาน สั่งconveyor เคลื่อที่ไปข้างหน้า" OR "ปุ่มClear",
                           PV := 1);
   "IEC_Counter_0_DB_154".CTUD(CU := ("Expected/Value_All".V = "Expected/Value_All".Expected_128) AND NOT "M128",
                           CD := "IEC_Counter_0_DB_1200".Q AND ("Barcode128" > 0) AND "ปุ่มยืนยันหน้า Screen",
                           PV := 5,
                           CV => "Barcode128");
   "M128" := "IEC_Counter_0_DB_154".QU;
   "IEC_Counter_0_DB_1201".CTU(CU := "ยา 129" = 1,
                           R := "Stepper Motor ทำงาน สั่งconveyor เคลื่อที่ไปข้างหน้า" OR "ปุ่มClear",
                           PV := 1);
   "IEC_Counter_0_DB_155".CTUD(CU := ("Expected/Value_All".V = "Expected/Value_All".Expected_129) AND NOT "M129",
                           CD := "IEC_Counter_0_DB_1201".Q AND ("Barcode129" > 0) AND "ปุ่มยืนยันหน้า Screen",
                           PV := 5,
                           CV => "Barcode129");
   "M129" := "IEC_Counter_0_DB_155".QU;
   "IEC_Counter_0_DB_1202".CTU(CU := "ยา 130" = 1,
                           R := "Stepper Motor ทำงาน สั่งconveyor เคลื่อที่ไปข้างหน้า" OR "ปุ่มClear",
                           PV := 1);
   "IEC_Counter_0_DB_156".CTUD(CU := ("Expected/Value_All".V = "Expected/Value_All".Expected_130) AND NOT "M130",
                           CD := "IEC_Counter_0_DB_1202".Q AND ("Barcode130" > 0) AND "ปุ่มยืนยันหน้า Screen",
                           PV := 5,
                           CV => "Barcode130");
   "M130" := "IEC_Counter_0_DB_156".QU;
   "IEC_Counter_0_DB_1203".CTU(CU := "ยา 131" = 1,
                           R := "Stepper Motor ทำงาน สั่งconveyor เคลื่อที่ไปข้างหน้า" OR "ปุ่มClear",
                           PV := 1);
   "IEC_Counter_0_DB_157".CTUD(CU := ("Expected/Value_All".V = "Expected/Value_All".Expected_131) AND NOT "M131",
                           CD := "IEC_Counter_0_DB_1203".Q AND ("Barcode131" > 0) AND "ปุ่มยืนยันหน้า Screen",
                           PV := 5,
                           CV => "Barcode131");
   "M131" := "IEC_Counter_0_DB_157".QU;
   "IEC_Counter_0_DB_1204".CTU(CU := "ยา 132" = 1,
                           R := "Stepper Motor ทำงาน สั่งconveyor เคลื่อที่ไปข้างหน้า" OR "ปุ่มClear",
                           PV := 1);
   "IEC_Counter_0_DB_158".CTUD(CU := ("Expected/Value_All".V = "Expected/Value_All".Expected_132) AND NOT "M132",
                           CD := "IEC_Counter_0_DB_1204".Q AND ("Barcode132" > 0) AND "ปุ่มยืนยันหน้า Screen",
                           PV := 5,
                           CV => "Barcode132");
   "M132" := "IEC_Counter_0_DB_158".QU;
   "IEC_Counter_0_DB_1205".CTU(CU := "ยา 133" = 1,
                           R := "Stepper Motor ทำงาน สั่งconveyor เคลื่อที่ไปข้างหน้า" OR "ปุ่มClear",
                           PV := 1);
   "IEC_Counter_0_DB_159".CTUD(CU := ("Expected/Value_All".V = "Expected/Value_All".Expected_133) AND NOT "M133",
                           CD := "IEC_Counter_0_DB_1205".Q AND ("Barcode133" > 0) AND "ปุ่มยืนยันหน้า Screen",
                           PV := 5,
                           CV => "Barcode133");
   "M133" := "IEC_Counter_0_DB_159".QU;
   "IEC_Counter_0_DB_1206".CTU(CU := "ยา 134" = 1,
                           R := "Stepper Motor ทำงาน สั่งconveyor เคลื่อที่ไปข้างหน้า" OR "ปุ่มClear",
                           PV := 1);
   "IEC_Counter_0_DB_160".CTUD(CU := ("Expected/Value_All".V = "Expected/Value_All".Expected_134) AND NOT "M134",
                           CD := "IEC_Counter_0_DB_1206".Q AND ("Barcode134" > 0) AND "ปุ่มยืนยันหน้า Screen",
                           PV := 5,
                           CV => "Barcode134");
   "M134" := "IEC_Counter_0_DB_160".QU;
   "IEC_Counter_0_DB_1207".CTU(CU := "ยา 135" = 1,
                           R := "Stepper Motor ทำงาน สั่งconveyor เคลื่อที่ไปข้างหน้า" OR "ปุ่มClear",
                           PV := 1);
   "IEC_Counter_0_DB_161".CTUD(CU := ("Expected/Value_All".V = "Expected/Value_All".Expected_135) AND NOT "M135",
                           CD := "IEC_Counter_0_DB_1207".Q AND ("Barcode135" > 0) AND "ปุ่มยืนยันหน้า Screen",
                           PV := 5,
                           CV => "Barcode135");
   "M135" := "IEC_Counter_0_DB_161".QU;
   "IEC_Counter_0_DB_1208".CTU(CU := "ยา 136" = 1,
                           R := "Stepper Motor ทำงาน สั่งconveyor เคลื่อที่ไปข้างหน้า" OR "ปุ่มClear",
                           PV := 1);
   "IEC_Counter_0_DB_162".CTUD(CU := ("Expected/Value_All".V = "Expected/Value_All".Expected_136) AND NOT "M136",
                           CD := "IEC_Counter_0_DB_1208".Q AND ("Barcode136" > 0) AND "ปุ่มยืนยันหน้า Screen",
                           PV := 5,
                           CV => "Barcode136");
   "M136" := "IEC_Counter_0_DB_162".QU;
   "IEC_Counter_0_DB_1209".CTU(CU := "ยา 137" = 1,
                           R := "Stepper Motor ทำงาน สั่งconveyor เคลื่อที่ไปข้างหน้า" OR "ปุ่มClear",
                           PV := 1);
   "IEC_Counter_0_DB_163".CTUD(CU := ("Expected/Value_All".V = "Expected/Value_All".Expected_137) AND NOT "M137",
                           CD := "IEC_Counter_0_DB_1209".Q AND ("Barcode137" > 0) AND "ปุ่มยืนยันหน้า Screen",
                           PV := 5,
                           CV => "Barcode137");
   "M137" := "IEC_Counter_0_DB_163".QU;
   "IEC_Counter_0_DB_1210".CTU(CU := "ยา 138" = 1,
                           R := "Stepper Motor ทำงาน สั่งconveyor เคลื่อที่ไปข้างหน้า" OR "ปุ่มClear",
                           PV := 1);
   "IEC_Counter_0_DB_164".CTUD(CU := ("Expected/Value_All".V = "Expected/Value_All".Expected_138) AND NOT "M138",
                           CD := "IEC_Counter_0_DB_1210".Q AND ("Barcode138" > 0) AND "ปุ่มยืนยันหน้า Screen",
                           PV := 5,
                           CV => "Barcode138");
   "M138" := "IEC_Counter_0_DB_164".QU;
   "IEC_Counter_0_DB_1211".CTU(CU := "ยา 139" = 1,
                           R := "Stepper Motor ทำงาน สั่งconveyor เคลื่อที่ไปข้างหน้า" OR "ปุ่มClear",
                           PV := 1);
   "IEC_Counter_0_DB_165".CTUD(CU := ("Expected/Value_All".V = "Expected/Value_All".Expected_139) AND NOT "M139",
                           CD := "IEC_Counter_0_DB_1211".Q AND ("Barcode139" > 0) AND "ปุ่มยืนยันหน้า Screen",
                           PV := 5,
                           CV => "Barcode139");
   "M139" := "IEC_Counter_0_DB_165".QU;
   "IEC_Counter_0_DB_1212".CTU(CU := "ยา 140" = 1,
                           R := "Stepper Motor ทำงาน สั่งconveyor เคลื่อที่ไปข้างหน้า" OR "ปุ่มClear",
                           PV := 1);
   "IEC_Counter_0_DB_166".CTUD(CU := ("Expected/Value_All".V = "Expected/Value_All".Expected_140) AND NOT "M140",
                           CD := "IEC_Counter_0_DB_1212".Q AND ("Barcode140" > 0) AND "ปุ่มยืนยันหน้า Screen",
                           PV := 5,
                           CV => "Barcode140");
   "M140" := "IEC_Counter_0_DB_166".QU;
END_REGION

REGION Network 8
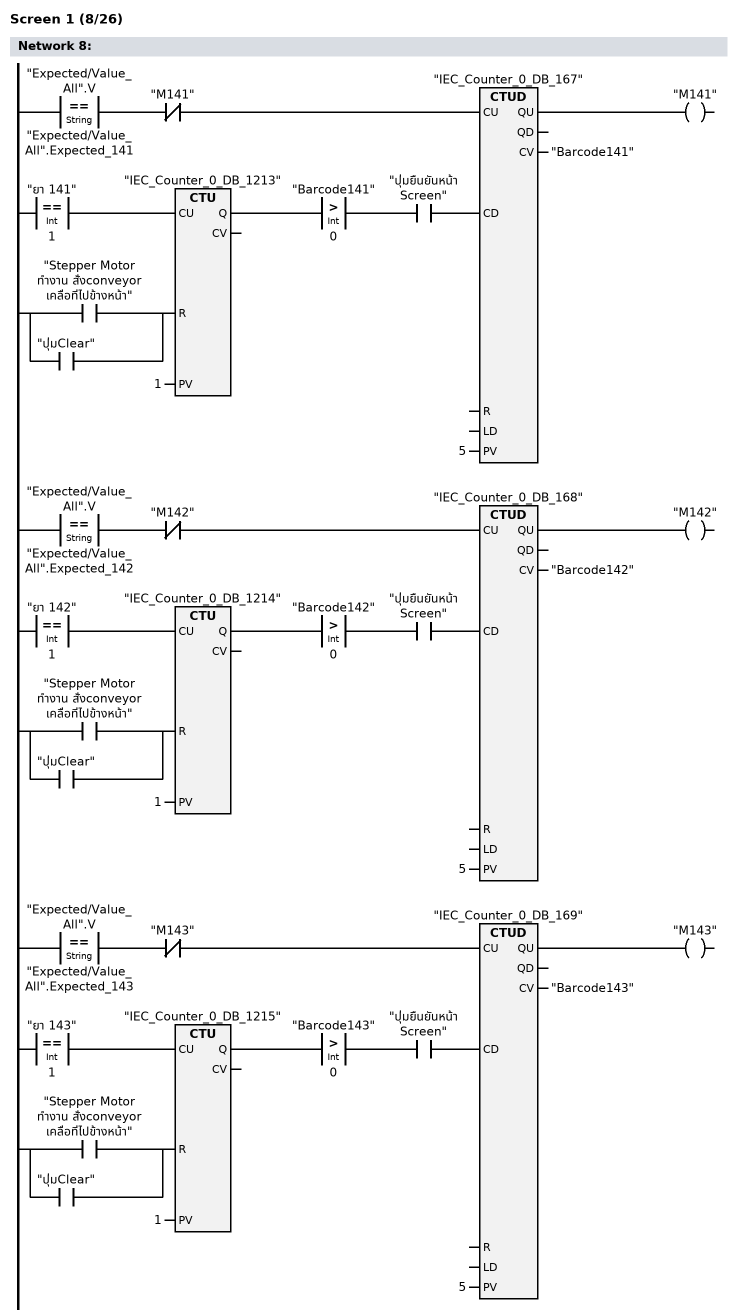
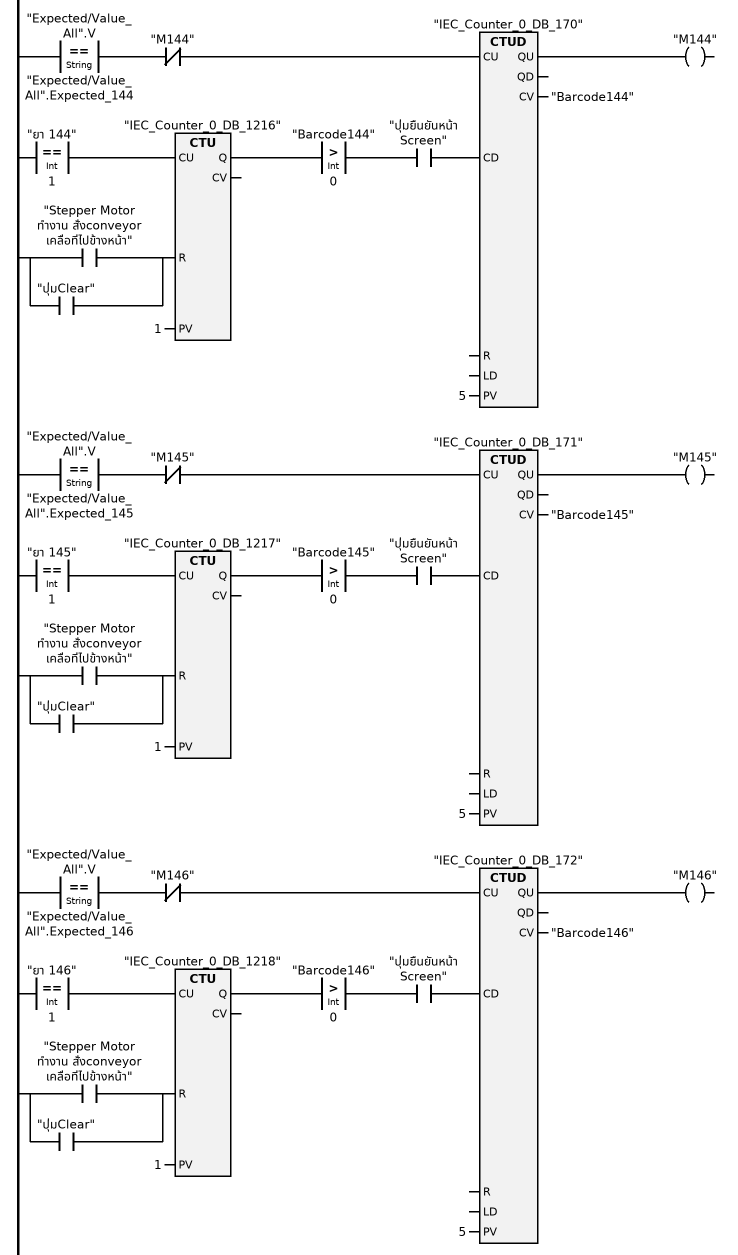
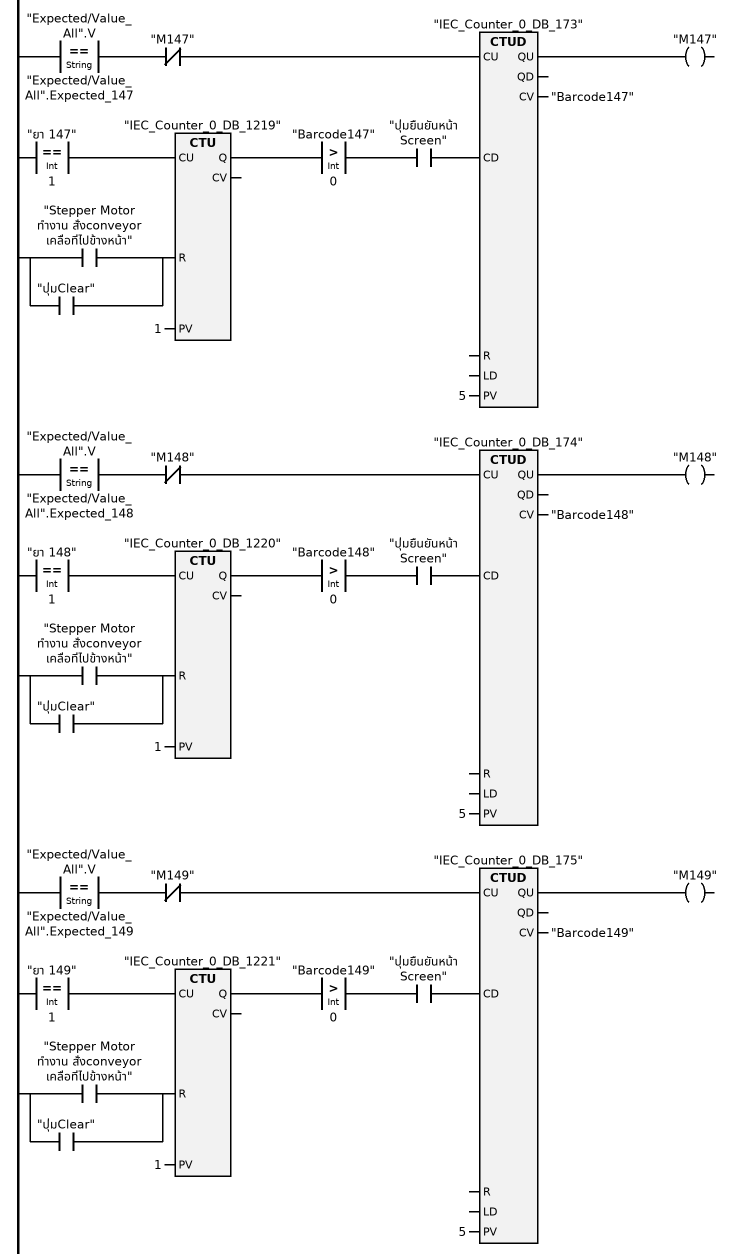
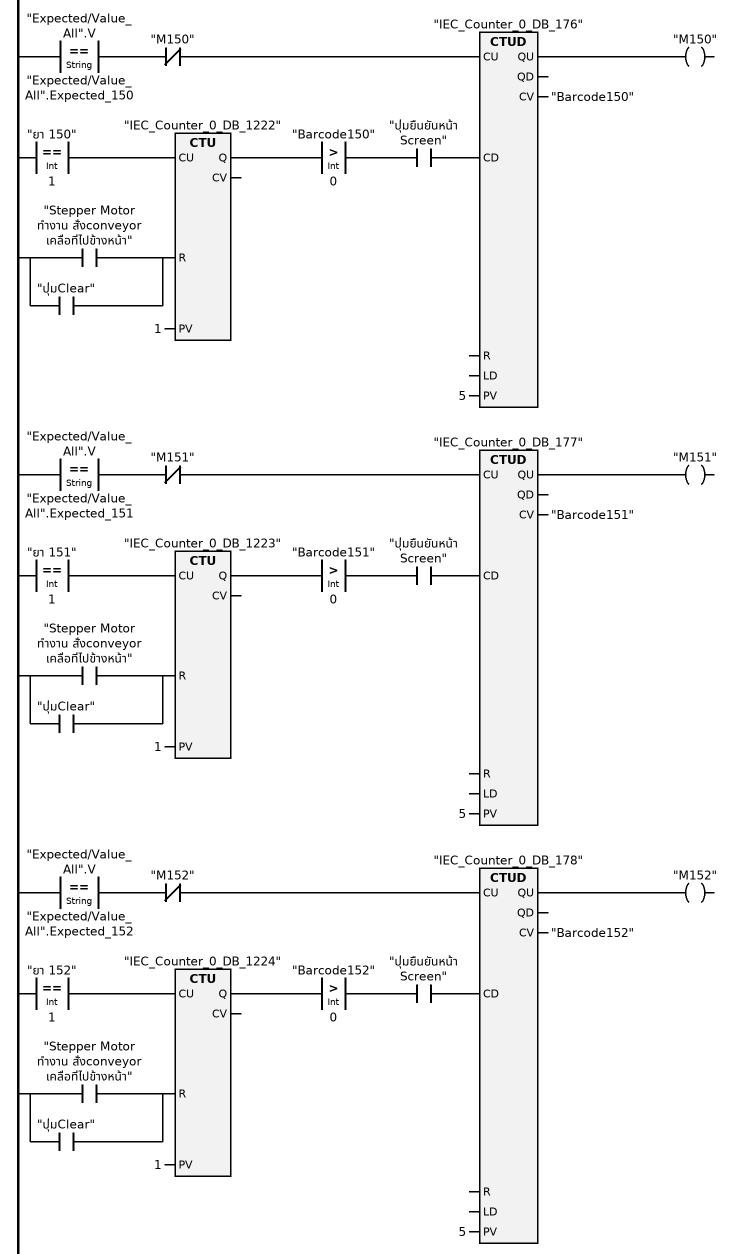
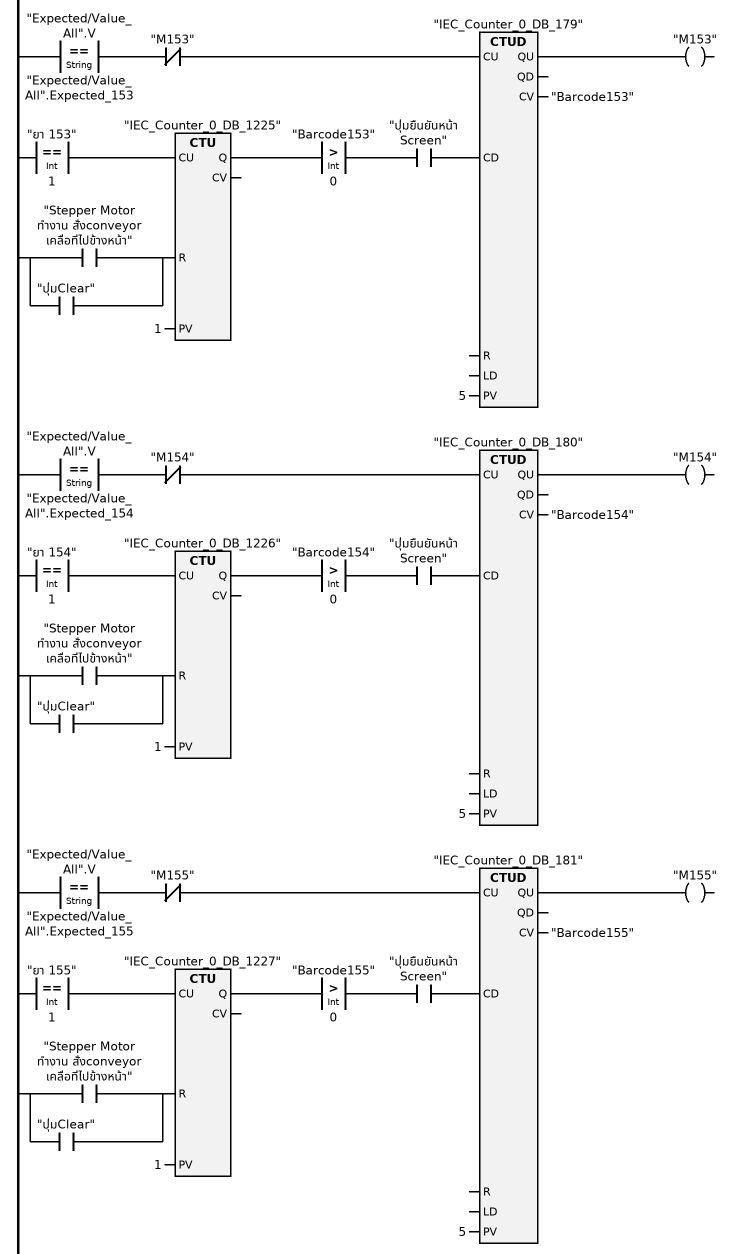
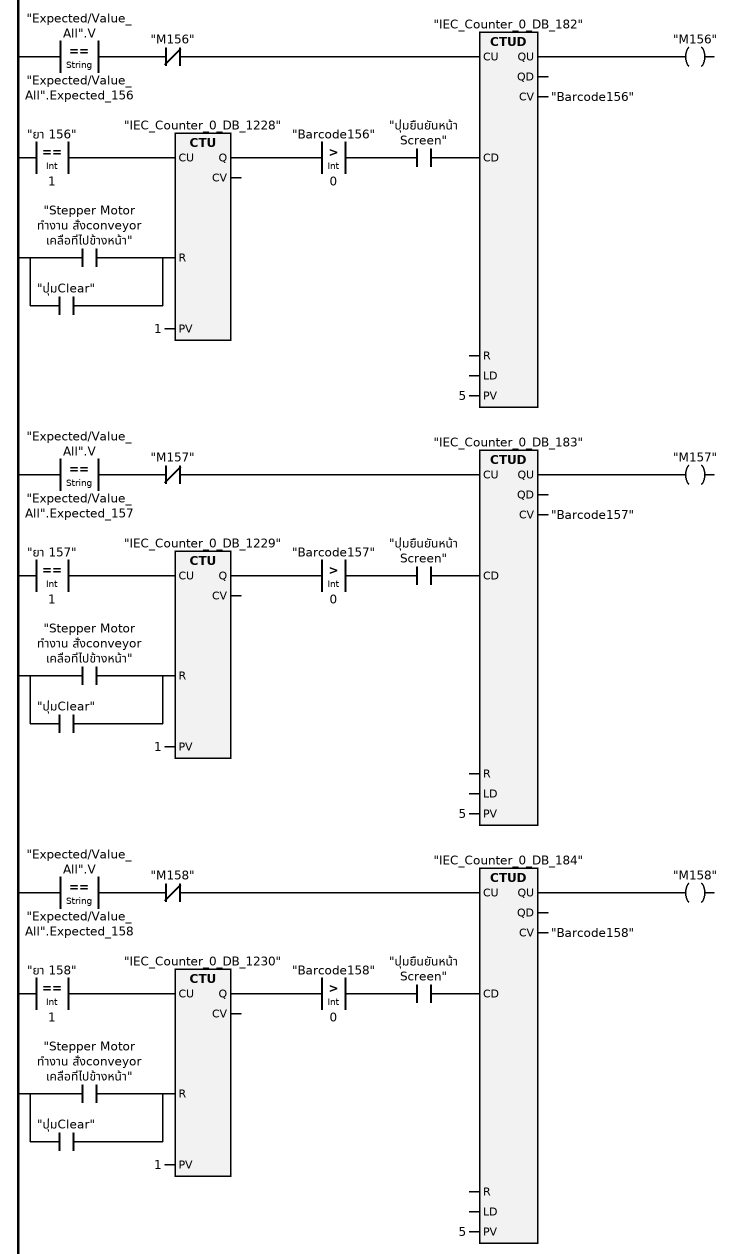
